(* IEC 61131-3 sources: rusty/tests/lit/cfc/connectors/chain, 1 file *)

(* ---- main.st ---- *)
FUNCTION main : DINT
    chain.foo := 7;
    chain();
    // CHECK: bar = 7
    printf('bar = %d$N', chain.bar);
END_FUNCTION
